SUBAPPLICATION logiBUS_PI_Speed_OPC (* logiBUS_PI Frequenz -> PT1-Filter -> SCALE/RASTER, Filterzeit/DerivK INI-persistiert, alles per OPC-UA (ohne VT) *)
  (* Standard: 61499-2; Description: Copyright (c) 2026 Meisterschulen am Ostbahnhof This program and the accompanying materials are made available under the terms of the Eclipse Public License 2.0 which is available at https://www.eclipse.org/legal/epl-2.0/ SPDX-License-Identifier: EPL-2.0 *)
  (* Version 1.0, 2026-10-28, Franz Höpfinger, Meisterschulen am Ostbahnhof, Kopie von MyLib::sys::logiBUS_PI_Speed_Publish_OPC ohne VT, fuer Stationen ohne VT (keine isobus_UT-Libs). FilterTimeS/DerivK -> MyLib::sys::OPC_TO_AR2_OUT, stObjFilterTimeS/stObjDerivK entfallen. Logik, INI-Keys und Defaults unveraendert. *)
  PACKAGE MyLib::sys;
  IMPORT logiBUS::io::PI::logiBUS_PI;
  IMPORT logiBUS::io::PI::logiBUS_PI_S;
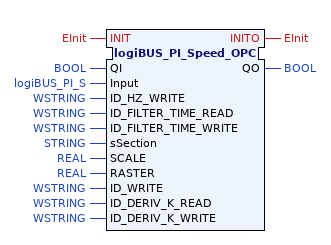
  EVENT_INPUT
    INIT : EInit; (* Initialization Request *)
  END_EVENT
  EVENT_OUTPUT
    INITO : EInit; (* Initialization Confirm *)
  END_EVENT
  VAR_INPUT
    QI : BOOL := TRUE; (* Quality Input - TRUE to enable service *)
    Input : logiBUS::io::PI::logiBUS_PI_S := logiBUS_PI::Invalid; (* Identify the Input PulseInput_I1..I9 *)
    ID_HZ_WRITE : WSTRING; (* Frequenz-Publish-Adresse (REAL Hz, ACTION=PUBLISH), lokal auf dieser Station - nur Dashboard/Diagnose, keine andere Station soll dies remote abonnieren (LOC-Scope) *)
    ID_FILTER_TIME_READ : WSTRING; (* Remote-Subscribe-Adresse (REAL Sekunden, ACTION=SUBSCRIBE) fuer Web-Override der Filterzeit *)
    ID_FILTER_TIME_WRITE : WSTRING; (* Lokale Echo/Re-Publish-Adresse (REAL Sekunden, ACTION=PUBLISH) der aktuellen Filterzeit *)
    sSection : STRING; (* INI settings.ini Section fuer die persistierte Filterzeit (eindeutig pro Sensor-Instanz) *)
    SCALE : REAL; (* Skalierungsfaktor Hz -> physikalische Einheit (z.B. 3.6/53 fuer km/h, 60.0 fuer U/min bei 1 Impuls/Umdrehung) *)
    RASTER : REAL := 0.001; (* Rundungsraster des FERTIGEN physikalischen Werts (nach SCALE), in der Anzeigeeinheit (z.B. 0.125 fuer U/min, 0.1 fuer km/h) - Platzhalter-Default 0.001 (praktisch kein Runden) *)
    ID_WRITE : WSTRING; (* Publish-Adresse des umgerechneten physikalischen Endwerts (REAL, ACTION=PUBLISH) - das ist die Adresse, die andere Stationen remote abonnieren (M2M-Scope) *)
    ID_DERIV_K_READ : WSTRING; (* Remote-Subscribe-Adresse (REAL, ACTION=SUBSCRIBE) fuer Web-Override von FT_DERIV_10_AR.K *)
    ID_DERIV_K_WRITE : WSTRING; (* Lokale Echo/Re-Publish-Adresse (REAL, ACTION=PUBLISH) des aktuellen FT_DERIV_10_AR.K *)
  END_VAR
  VAR_OUTPUT
    QO : BOOL; (* Quality Output - TRUE if service executed successfully *)
  END_VAR
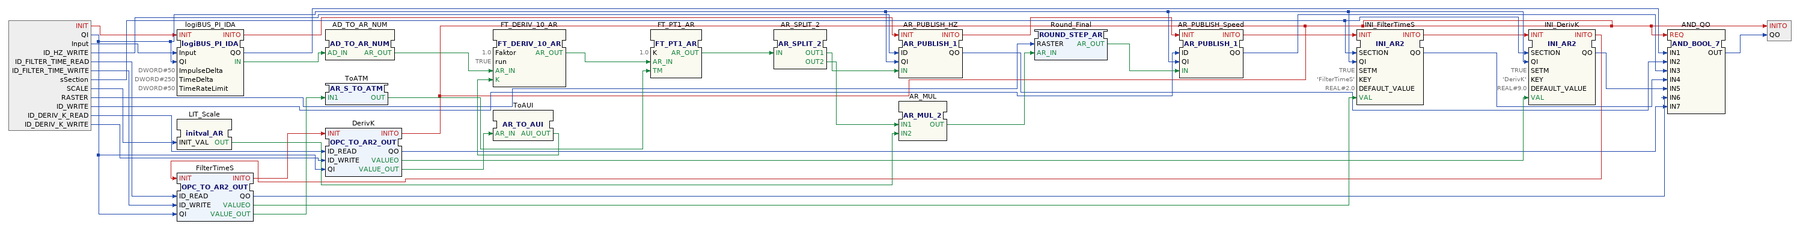
  FBS
    logiBUS_PI_IDA : logiBUS::io::PI::logiBUS_PI_IDA(ImpulseDelta := DWORD#50, TimeDelta := DWORD#250, TimeRateLimit := DWORD#50);
    AD_TO_AR_NUM : adapter::conversion::unidirectional::AD_TO_AR_NUM;
    FT_DERIV_10_AR : OSCAT_adapter::Control::FT_DERIV_10_AR(Faktor := 1.0, run := TRUE);
    FT_PT1_AR : OSCAT_adapter::Control::FT_PT1_AR(K := 1.0);
    AR_SPLIT_2 : adapter::events::unidirectional::AR_SPLIT_2;
    AR_PUBLISH_HZ : adapter::net::AR_PUBLISH_1;
    LIT_Scale : adapter::types::unidirectional::AR::initval::initval_AR;
    AR_MUL : adapter::iec61131::arithmetic::AR_MUL_2;
    AR_PUBLISH_Speed : adapter::net::AR_PUBLISH_1;
    INI_FilterTimeS : eclipse4diac::storage::INI_AR2(SETM := TRUE, KEY := 'FilterTimeS', DEFAULT_VALUE := REAL#2.0);
    INI_DerivK : eclipse4diac::storage::INI_AR2(SETM := TRUE, KEY := 'DerivK', DEFAULT_VALUE := REAL#9.0);
    ToAUI : adapter::conversion::unidirectional::AR_TO_AUI;
    AND_QO : iec61131::booleanOperators::AND_BOOL_7;
  END_FBS
  SUBAPPS
    Round_Final : OSCAT_adapter::Mathematical::ROUND_STEP_AR;
    FilterTimeS : MyLib::sys::OPC_TO_AR2_OUT;
    ToATM : MyLib::sys::AR_S_TO_ATM;
    DerivK : MyLib::sys::OPC_TO_AR2_OUT;
  END_SUBAPPS
  EVENT_CONNECTIONS
    INIT TO logiBUS_PI_IDA.INIT;
    logiBUS_PI_IDA.INITO TO AR_PUBLISH_HZ.INIT;
    AR_PUBLISH_HZ.INITO TO AR_PUBLISH_Speed.INIT;
    AR_PUBLISH_Speed.INITO TO INI_FilterTimeS.INIT;
    INI_FilterTimeS.INITO TO INI_DerivK.INIT;
    INI_DerivK.INITO TO FilterTimeS.INIT;
    FilterTimeS.INITO TO DerivK.INIT;
    DerivK.INITO TO INITO;
    DerivK.INITO TO AND_QO.REQ;
  END_CONNECTIONS
  DATA_CONNECTIONS
    Input TO logiBUS_PI_IDA.Input;
    ID_HZ_WRITE TO AR_PUBLISH_HZ.ID;
    ID_FILTER_TIME_READ TO FilterTimeS.ID_READ;
    ID_FILTER_TIME_WRITE TO FilterTimeS.ID_WRITE;
    sSection TO INI_FilterTimeS.SECTION;
    SCALE TO LIT_Scale.INIT_VAL;
    RASTER TO Round_Final.RASTER;
    ID_WRITE TO AR_PUBLISH_Speed.ID;
    ID_DERIV_K_READ TO DerivK.ID_READ;
    ID_DERIV_K_WRITE TO DerivK.ID_WRITE;
    sSection TO INI_DerivK.SECTION;
    QI TO logiBUS_PI_IDA.QI;
    QI TO AR_PUBLISH_HZ.QI;
    QI TO AR_PUBLISH_Speed.QI;
    QI TO INI_FilterTimeS.QI;
    QI TO INI_DerivK.QI;
    logiBUS_PI_IDA.QO TO AND_QO.IN1;
    AR_PUBLISH_HZ.QO TO AND_QO.IN2;
    AR_PUBLISH_Speed.QO TO AND_QO.IN3;
    INI_FilterTimeS.QO TO AND_QO.IN4;
    INI_DerivK.QO TO AND_QO.IN5;
    AND_QO.OUT TO QO;
    QI TO FilterTimeS.QI;
    QI TO DerivK.QI;
    FilterTimeS.QO TO AND_QO.IN6;
    DerivK.QO TO AND_QO.IN7;
  END_CONNECTIONS
  ADAPTER_CONNECTIONS
    logiBUS_PI_IDA.IN TO AD_TO_AR_NUM.AD_IN;
    AD_TO_AR_NUM.AR_OUT TO FT_DERIV_10_AR.AR_IN;
    FT_DERIV_10_AR.AR_OUT TO FT_PT1_AR.AR_IN;
    FilterTimeS.VALUEO TO INI_FilterTimeS.VAL;
    FilterTimeS.VALUE_OUT TO ToATM.IN1;
    ToATM.OUT TO FT_PT1_AR.TM;
    FT_PT1_AR.AR_OUT TO AR_SPLIT_2.IN;
    AR_SPLIT_2.OUT1 TO AR_PUBLISH_HZ.IN;
    AR_SPLIT_2.OUT2 TO AR_MUL.IN1;
    LIT_Scale.OUT TO AR_MUL.IN2;
    AR_MUL.OUT TO Round_Final.AR_IN;
    Round_Final.AR_OUT TO AR_PUBLISH_Speed.IN;
    DerivK.VALUEO TO INI_DerivK.VAL;
    DerivK.VALUE_OUT TO ToAUI.AR_IN;
    ToAUI.AUI_OUT TO FT_DERIV_10_AR.K;
  END_CONNECTIONS
END_SUBAPPLICATION
